// TIA Portal V21 export
// export: Created 2026-11-11T00:47:41.1020194Z, ExportSetting WithDefaults, DisplayName Totally Integrated Automation Portal, DisplayVersion V21 Update 3, DisplayName STEP 7 Professional, DisplayVersion V21 Update 3, DisplayName STEP 7 Safety, DisplayVersion V21, DisplayName Tech WebApplication, DisplayVersion V21, DisplayName WinCC Basic/Comfort/Advanced, DisplayVersion V21 Update 3, DisplayName WinCC Unified, DisplayVersion V21 Update 3
FUNCTION_BLOCK "FB_Fbd_ex155"   // FB163, FBD
{ S7_Optimized_Access := 'TRUE' }
VERSION : 0.1
// stored: AutoNumber true, IsIECCheckEnabled false, IsRetainMemResEnabled false, MemoryReserve 100, SetENOAutomatically false, UDAEnableTagReadback false
   VAR_INPUT
      v_addr : Variant;
   END_VAR
   VAR_OUTPUT
      v_ret_val : Int;
      v_laddr : HW_IO;
   END_VAR
BEGIN

REGION Network 1: IO2MOD - Determine hardware identifier from an IO address
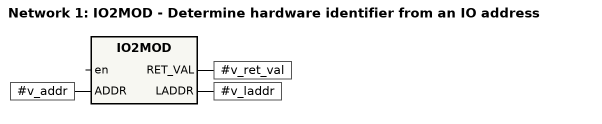
   #v_ret_val := IO2MOD(ADDR := #v_addr, LADDR => #v_laddr);
END_REGION
END_FUNCTION_BLOCK
